(* IEC 61131-3 sources: Elmo_Master/Lasal_PRG/MotionTCPDemo/Class/UDPTransmission, 1 file *)

(* ---- UDPTransmission.st ---- *)
#define IP_ADDR_MIN_LEN         7
#define IP_ADDR_MAX_LEN         15

(*!
<Class
	Name               = "UDPTransmission"
	Revision           = "0.0"
	RealtimeTask       = "true"
	CyclicTask         = "true"
	BackgroundTask     = "false"
	Sigmatek           = "false"
	OSInterface        = "false"
	HighPriority       = "false"
	Automatic          = "false"
	UpdateMode         = "Prescan"
	SharedCommandTable = "true"
	Objectsize         = "(536,120)">
	<Channels>
		<Server Name="Dbg_RecMsg" Visualized="false" Initialize="false" WriteProtected="true" Retentive="false"/>
		<Server Name="Dbg_SendMsg" Visualized="false" Initialize="false" WriteProtected="true" Retentive="false"/>
		<Server Name="RecMsg32" Visualized="false" Initialize="false" WriteProtected="true" Retentive="false"/>
		<Server Name="TransError" Visualized="false" Initialize="false" WriteProtected="true" Retentive="false"/>
		<Server Name="TransState" Visualized="false" Initialize="false" WriteProtected="true" Retentive="false"/>
		<Client Name="IPAddr" Required="true" Internal="false"/>
		<Client Name="Port" Required="true" Internal="false"/>
	</Channels>
	<Network Name="UDPTransmission">
		<!-- List of Components in this network -->
		<Components>
			<Object
				Name       = "_base"
				Class      = "_UDPTransceiverInterface"
				Position   = "(218,120)"
				Visualized = "true"
				Remotely   = "true">
				<Channels>
					<Server Name="ClassSvr"/>
					<Server Name="ErrorCode"/>
					<Server Name="ErrorMessage"/>
					<Server Name="ErrorState"/>
					<Server Name="State"/>
					<Client Name="_UDPTransceiver"/>
				</Channels>
			</Object>
		</Components>
		<Comments>
		</Comments>
		<!-- List of Connections in this network -->
		<Connections>
			<Connection Source="this.ClassSvr" Destination="_base.ClassSvr" Vertices="(942,210),(770,210),"/>
			<Connection Source="this.State" Destination="_base.State" Vertices="(942,270),(770,270),"/>
			<Connection Source="this.ErrorState" Destination="_base.ErrorState" Vertices="(942,330),(770,330),"/>
			<Connection Source="this.ErrorMessage" Destination="_base.ErrorMessage" Vertices="(942,390),(770,390),"/>
			<Connection Source="this.ErrorCode" Destination="_base.ErrorCode" Vertices="(942,450),(770,450),"/>
			<Connection Source="_base._UDPTransceiver" Destination="this._UDPTransceiver" Vertices="(218,210),(38,210),"/>
		</Connections>
		<!-- Headerfiles -->
		<Options>
		</Options>
	</Network>
</Class>
*)
#pragma using _UDPTransceiverInterface

UDPTransmission : CLASS
: _UDPTransceiverInterface
	TYPE
	  t_e_TransmissionState :  //! <Type Public="true" Name="t_e_TransmissionState"/>
	  (
	    TS_CheckPara,
	    TS_AddSocket,
	    TS_CheckSocket,
	    TS_BindRecSocket,
	    TS_SendData,
	    TS_Error
	  )$UDINT;
#pragma pack(push, 1)
	  t_s_BrakeDataSend : STRUCT
	    ActForce : DINT;
	    ActPos : DINT;
	  END_STRUCT;
#pragma pack(pop)
	END_TYPE
  //Servers:
	TransState 	: SvrCh_t_e_TransmissionState_PTofCls_UDPTransmission;
	TransError 	: SvrCh_DINT;
	Dbg_SendMsg 	: SvrCh_DINT;
	Dbg_RecMsg 	: SvrCh_DINT;
	RecMsg32 	: SvrCh_DINT;
  //Clients:
	IPAddr 	: CltChCmd_String;
	Port 	: CltCh_DINT;
  //Variables:
		BrakeData 	: t_s_BrakeDataSend;
		IPDest : ARRAY [0..IP_ADDR_MAX_LEN] OF CHAR;

		udIPDest 	: UDINT;
		IPSrc : ARRAY [0..IP_ADDR_MAX_LEN] OF CHAR;

		udIPSrc 	: UDINT;
  //Functions:

	FUNCTION VIRTUAL GLOBAL CyWork
		VAR_INPUT
			EAX 	: UDINT;
		END_VAR
		VAR_OUTPUT
			state (EAX) 	: UDINT;
		END_VAR;

	FUNCTION VIRTUAL GLOBAL RtWork
		VAR_INPUT
			EAX 	: UDINT;
		END_VAR
		VAR_OUTPUT
			state (EAX) 	: UDINT;
		END_VAR;
				//! <Function Comment="function is called when a complete package has been received" Name="Response"/>
	FUNCTION VIRTUAL GLOBAL Response
		VAR_INPUT
			pData 	: ^void;			//! <Variable Comment="pointer to received data" Name="Response.pData"/>
			udsize 	: UDINT;			//! <Variable Comment="size of received package" Name="Response.udsize"/>
			SourceIP 	: UDINT;
			SourcePort 	: UDINT;
		END_VAR;
  //Tables:
	FUNCTION @STD
		VAR_OUTPUT
			ret_code	: CONFSTATES;
		END_VAR;
	FUNCTION GLOBAL TAB @CT_;
END_CLASS;

#pragma usingLtd String

FUNCTION VIRTUAL GLOBAL UDPTransmission::RtWork
	VAR_INPUT
		EAX 	: UDINT;
	END_VAR
	VAR_OUTPUT
		state (EAX) 	: UDINT;
	END_VAR
  VAR
	tmpLen : UDINT;
  END_VAR

  //**************************************************************************************
  //**************************************************************************************
  case TransState of
    //************************************************************************************
	TS_CheckPara: // check if ip address and port are meaningful
    //************************************************************************************
     IPAddr.TxtToAscii();
     tmpLen := IPAddr.TxtLen();
     if tmpLen < IP_ADDR_MIN_LEN | tmpLen > IP_ADDR_MAX_LEN then
      TransError := -1;
      TransState := TS_Error;
     end_if;

     IPAddr.TxtGet(pdst:=#IPDest[0], dstsize:=sizeof(IPDest));

     udIPDest := _UDPTransceiver.ConvertStrToUdint(pIpAddress:=#IPDest[0]);

     Port := Port.Read();

     TransState := TS_AddSocket;

    //************************************************************************************
	TS_AddSocket: // trigger opening of socked
    //************************************************************************************

      AddSocket();
      TransState := TS_CheckSocket;

    //************************************************************************************
	TS_CheckSocket: // check if socket is open
    //************************************************************************************
      if IsOpen() then

        TransState := TS_SendData;
      end_if;
    //************************************************************************************
	TS_BindRecSocket: // check if socket is open
    //************************************************************************************

      if GetIpInfo(pIpInfo:=#udIPSrc, dPara:=IP_OPT_ADDR, dInterface:=1) then
        _UDPTransceiver.ConvertUdintToStr(pIpAddress:=#IPSrc[0], udLen:=sizeof(IPSrc), udIpAddress:=udIPSrc);

        if BindSocket(pIpAddress:=#IPSrc[0], udPort:=to_udint(Port.Read())) <> 0 then
          TransError := -2;
        end_if;
      else
        TransError := -3;
      end_if;

      TransState := TS_SendData;

    //************************************************************************************
	TS_SendData:
    //************************************************************************************

    //************************************************************************************
	TS_Error:
    //************************************************************************************
  end_case;
  //**************************************************************************************
  //**************************************************************************************

	state := READY;

END_FUNCTION

FUNCTION VIRTUAL GLOBAL UDPTransmission::CyWork
	VAR_INPUT
		EAX 	: UDINT;
	END_VAR
	VAR_OUTPUT
		state (EAX) 	: UDINT;
	END_VAR
  VAR
	tmpLen : UDINT;
  END_VAR

  //**************************************************************************************
  //**************************************************************************************
  case TransState of
    //************************************************************************************
	TS_CheckPara: // check if ip address and port are meaningful
    //************************************************************************************
     IPAddr.TxtToAscii();
     tmpLen := IPAddr.TxtLen();
     if tmpLen < IP_ADDR_MIN_LEN | tmpLen > IP_ADDR_MAX_LEN then
      TransError := -1;
      TransState := TS_Error;
     end_if;

     IPAddr.TxtGet(pdst:=#IPDest[0], dstsize:=16);

     udIPDest := _UDPTransceiver.ConvertStrToUdint(pIpAddress:=#IPDest[0]);

     Port := Port.Read();

     TransState := TS_AddSocket;

    //************************************************************************************
	TS_AddSocket: // trigger opening of socked
    //************************************************************************************

      AddSocket();

      TransState := TS_CheckSocket;

    //************************************************************************************
	TS_CheckSocket: // check if socket is open
    //************************************************************************************
      if IsOpen() then
        TransState := TS_BindRecSocket;
      end_if;

    //************************************************************************************
	TS_BindRecSocket: // check if socket is open
    //************************************************************************************
      if GetIpInfo(pIpInfo:=#udIPSrc, dPara:=IP_OPT_ADDR, dInterface:=1) = 0 then
        _UDPTransceiver.ConvertUdintToStr(pIpAddress:=#IPSrc[0], udLen:=sizeof(IPSrc), udIpAddress:=udIPSrc);

        if BindSocket(pIpAddress:=#IPSrc[0], udPort:=to_udint(Port.Read())) < 0 then
          TransError := -2;
        end_if;
      else
        TransError := -3;
      end_if;

      TransState := TS_SendData;

    //************************************************************************************
	TS_SendData:
    //************************************************************************************

    //************************************************************************************
	TS_Error:
    //************************************************************************************
  end_case;
  //**************************************************************************************
  //**************************************************************************************

	state := READY;

END_FUNCTION

FUNCTION VIRTUAL GLOBAL UDPTransmission::Response
	VAR_INPUT
		pData 	: ^void;
		udsize 	: UDINT;
		SourceIP 	: UDINT;
		SourcePort 	: UDINT;
	END_VAR

  if pData <> NIL & udsize > 0 then

    RecMsg32 := pData^$DINT;
    Dbg_RecMsg += 1;

  end_if;

END_FUNCTION
